TYPE "ST_ModelField"
VERSION : 0.1
   STRUCT
      "Name" : String[32];
      "Value" : String[64];
   END_STRUCT;
END_TYPE
